//One client of the Siemens simulator
TYPE ST_Sim_Client :
STRUCT
	nClient	: INT;					//0 = empty position
	eRecipe	: E_Anybus_RecipeType;
	eType	: E_Anybus_ClientType;
END_STRUCT
END_TYPE

(* stored: Version 1.1.0.1, ProductVersion 3.1.4026.20
   DUT ST_Sim_Client: Id {6c1f0a54-2b7e-4f0e-9d3a-1e5b7a90c103} *)
